ORGANIZATION_BLOCK "ProgramCycle"
TITLE = "Main Program Sweep (Cycle)"
{ S7_Optimized_Access := 'TRUE' }
VERSION : 0.1

BEGIN
    // Единственный вызов: всю работу делает оркестратор "ConveyorMain".
    // Слои вызываются внутри него в порядке: вход → логика → выход → ЧМИ.
    "ConveyorMain_DB"();
END_ORGANIZATION_BLOCK
